INTERFACE I_EtherCAT

PROPERTY inError : BOOL
GET
END_GET
END_PROPERTY

END_INTERFACE

(* stored: Version 1.1.0.1, ProductVersion 3.1.4024.12
   Itf I_EtherCAT: Id {56712762-1537-474d-beb1-103e887f2ab4}
   Property inError: Id {2234d776-9fe3-42a5-8a61-b133c29a043e}
   Get Get: Id {b5596eb6-36db-40ba-aa0a-f2287b7ce024} *)
